Universal Robots PolyScope program: SplitTest.urp

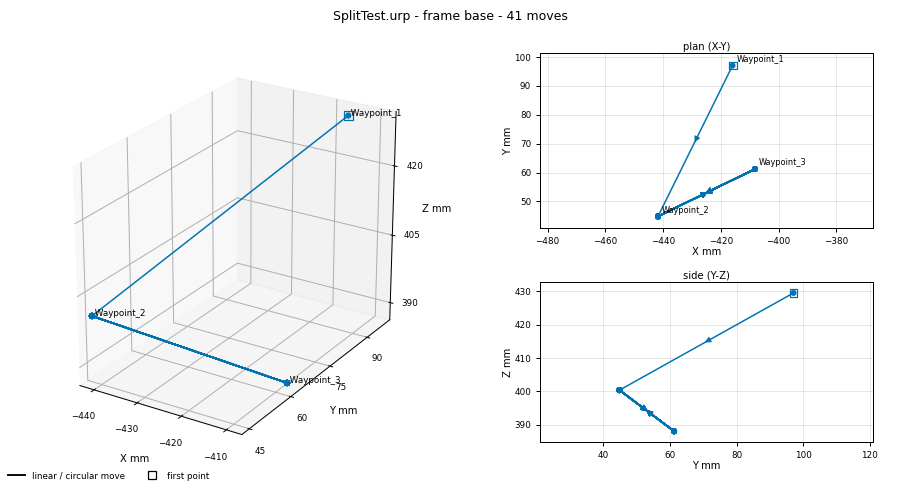
[picture p0: tool path of SplitTest.urp in frame base, 41 of 41 moves have a stored position in this frame; points joined in program order, loops and branches not executed]
Program SplitTest (createdIn=3.0.0 lastSavedIn=3.0.0 directory=/programs installation=default)
Robot Program (runOnlyOnce=true motionType=MoveJ speed=1.047198 acceleration=1.396263 useActiveTCP=false)
  'Program generated by VerticalBot Studio for UR5e on 25/10/2026 12:00:00'
  'Using nominal kinematics.'
  'Using Ref. Frame 2: p[0.100000, -0.050000, 0.020000, 0.000000, 0.000000, 0.523599]'
  'Using TCP Tool 1: p[0.010000, 0.000000, 0.120000, 0.000000, 0.261799, 0.000000]'
  Script: set_tcp(p[0.010000, 0.000000, 0.120000, 0.000000, 0.261799, 0.000000])
  Script: movej([-0.523599, -1.745329, 1.570796, -1.396263, -1.570796, 0.349066],1.20000,0.75000,0,0.0000)
  MoveJ speed 42.97 deg/s, acceleration 68.75 deg/s^2 (useActiveTCP=true)
    Waypoint Waypoint_1: TCP in base x=-415.957 y=97.082 z=429.557 mm, rx=-2.8465 ry=-1.036 rz=-0.3747 rad; joints [-30, -100, 90, -80, -90, 20] deg; flange x=-423.617 y=90.654 z=549.557 mm, rx=2.9521 ry=1.0745 rz=0 rad
  MoveL speed 200 mm/s, acceleration 1200 mm/s^2 (useActiveTCP=true)
    Waypoint Waypoint_2: TCP in base x=-441.769 y=44.852 z=400.392 mm, rx=-2.784 ry=-1.254 rz=-0.442 rad; joints [-22, -96, 90, -80, -90, 20] deg; flange x=-456.215 y=40.554 z=519.861 mm, rx=2.8233 ry=1.257 rz=0.075 rad
    Waypoint Waypoint_3: TCP in base x=-408.198 y=61.237 z=388.074 mm, rx=-2.843 ry=-1.1666 rz=-0.4658 rad; joints [-26, -100, 95, -80, -90, 20] deg; flange x=-424.78 y=58.869 z=507.319 mm, rx=2.8515 ry=1.1521 rz=0.0898 rad
    Waypoint Waypoint_4: TCP in base x=-441.769 y=44.852 z=400.392 mm, rx=-2.784 ry=-1.254 rz=-0.442 rad; joints [-22, -96, 90, -80, -90, 20] deg; flange x=-456.215 y=40.554 z=519.861 mm, rx=2.8233 ry=1.257 rz=0.075 rad
    Waypoint Waypoint_5: TCP in base x=-408.198 y=61.237 z=388.074 mm, rx=-2.843 ry=-1.1666 rz=-0.4658 rad; joints [-26, -100, 95, -80, -90, 20] deg; flange x=-424.78 y=58.869 z=507.319 mm, rx=2.8515 ry=1.1521 rz=0.0898 rad
    Waypoint Waypoint_6: TCP in base x=-441.769 y=44.852 z=400.392 mm, rx=-2.784 ry=-1.254 rz=-0.442 rad; joints [-22, -96, 90, -80, -90, 20] deg; flange x=-456.215 y=40.554 z=519.861 mm, rx=2.8233 ry=1.257 rz=0.075 rad
    Waypoint Waypoint_7: TCP in base x=-408.198 y=61.237 z=388.074 mm, rx=-2.843 ry=-1.1666 rz=-0.4658 rad; joints [-26, -100, 95, -80, -90, 20] deg; flange x=-424.78 y=58.869 z=507.319 mm, rx=2.8515 ry=1.1521 rz=0.0898 rad
    Waypoint Waypoint_8: TCP in base x=-441.769 y=44.852 z=400.392 mm, rx=-2.784 ry=-1.254 rz=-0.442 rad; joints [-22, -96, 90, -80, -90, 20] deg; flange x=-456.215 y=40.554 z=519.861 mm, rx=2.8233 ry=1.257 rz=0.075 rad
    Waypoint Waypoint_9: TCP in base x=-408.198 y=61.237 z=388.074 mm, rx=-2.843 ry=-1.1666 rz=-0.4658 rad; joints [-26, -100, 95, -80, -90, 20] deg; flange x=-424.78 y=58.869 z=507.319 mm, rx=2.8515 ry=1.1521 rz=0.0898 rad
    Waypoint Waypoint_10: TCP in base x=-441.769 y=44.852 z=400.392 mm, rx=-2.784 ry=-1.254 rz=-0.442 rad; joints [-22, -96, 90, -80, -90, 20] deg; flange x=-456.215 y=40.554 z=519.861 mm, rx=2.8233 ry=1.257 rz=0.075 rad
    Waypoint Waypoint_11: TCP in base x=-408.198 y=61.237 z=388.074 mm, rx=-2.843 ry=-1.1666 rz=-0.4658 rad; joints [-26, -100, 95, -80, -90, 20] deg; flange x=-424.78 y=58.869 z=507.319 mm, rx=2.8515 ry=1.1521 rz=0.0898 rad
    Waypoint Waypoint_12: TCP in base x=-441.769 y=44.852 z=400.392 mm, rx=-2.784 ry=-1.254 rz=-0.442 rad; joints [-22, -96, 90, -80, -90, 20] deg; flange x=-456.215 y=40.554 z=519.861 mm, rx=2.8233 ry=1.257 rz=0.075 rad
    Waypoint Waypoint_13: TCP in base x=-408.198 y=61.237 z=388.074 mm, rx=-2.843 ry=-1.1666 rz=-0.4658 rad; joints [-26, -100, 95, -80, -90, 20] deg; flange x=-424.78 y=58.869 z=507.319 mm, rx=2.8515 ry=1.1521 rz=0.0898 rad
    Waypoint Waypoint_14: TCP in base x=-441.769 y=44.852 z=400.392 mm, rx=-2.784 ry=-1.254 rz=-0.442 rad; joints [-22, -96, 90, -80, -90, 20] deg; flange x=-456.215 y=40.554 z=519.861 mm, rx=2.8233 ry=1.257 rz=0.075 rad
    Waypoint Waypoint_15: TCP in base x=-408.198 y=61.237 z=388.074 mm, rx=-2.843 ry=-1.1666 rz=-0.4658 rad; joints [-26, -100, 95, -80, -90, 20] deg; flange x=-424.78 y=58.869 z=507.319 mm, rx=2.8515 ry=1.1521 rz=0.0898 rad
    Waypoint Waypoint_16: TCP in base x=-441.769 y=44.852 z=400.392 mm, rx=-2.784 ry=-1.254 rz=-0.442 rad; joints [-22, -96, 90, -80, -90, 20] deg; flange x=-456.215 y=40.554 z=519.861 mm, rx=2.8233 ry=1.257 rz=0.075 rad
    Waypoint Waypoint_17: TCP in base x=-408.198 y=61.237 z=388.074 mm, rx=-2.843 ry=-1.1666 rz=-0.4658 rad; joints [-26, -100, 95, -80, -90, 20] deg; flange x=-424.78 y=58.869 z=507.319 mm, rx=2.8515 ry=1.1521 rz=0.0898 rad
    Waypoint Waypoint_18: TCP in base x=-441.769 y=44.852 z=400.392 mm, rx=-2.784 ry=-1.254 rz=-0.442 rad; joints [-22, -96, 90, -80, -90, 20] deg; flange x=-456.215 y=40.554 z=519.861 mm, rx=2.8233 ry=1.257 rz=0.075 rad
    Waypoint Waypoint_19: TCP in base x=-408.198 y=61.237 z=388.074 mm, rx=-2.843 ry=-1.1666 rz=-0.4658 rad; joints [-26, -100, 95, -80, -90, 20] deg; flange x=-424.78 y=58.869 z=507.319 mm, rx=2.8515 ry=1.1521 rz=0.0898 rad
    Waypoint Waypoint_20: TCP in base x=-441.769 y=44.852 z=400.392 mm, rx=-2.784 ry=-1.254 rz=-0.442 rad; joints [-22, -96, 90, -80, -90, 20] deg; flange x=-456.215 y=40.554 z=519.861 mm, rx=2.8233 ry=1.257 rz=0.075 rad
    Waypoint Waypoint_21: TCP in base x=-408.198 y=61.237 z=388.074 mm, rx=-2.843 ry=-1.1666 rz=-0.4658 rad; joints [-26, -100, 95, -80, -90, 20] deg; flange x=-424.78 y=58.869 z=507.319 mm, rx=2.8515 ry=1.1521 rz=0.0898 rad
    Waypoint Waypoint_22: TCP in base x=-441.769 y=44.852 z=400.392 mm, rx=-2.784 ry=-1.254 rz=-0.442 rad; joints [-22, -96, 90, -80, -90, 20] deg; flange x=-456.215 y=40.554 z=519.861 mm, rx=2.8233 ry=1.257 rz=0.075 rad
    Waypoint Waypoint_23: TCP in base x=-408.198 y=61.237 z=388.074 mm, rx=-2.843 ry=-1.1666 rz=-0.4658 rad; joints [-26, -100, 95, -80, -90, 20] deg; flange x=-424.78 y=58.869 z=507.319 mm, rx=2.8515 ry=1.1521 rz=0.0898 rad
    Waypoint Waypoint_24: TCP in base x=-441.769 y=44.852 z=400.392 mm, rx=-2.784 ry=-1.254 rz=-0.442 rad; joints [-22, -96, 90, -80, -90, 20] deg; flange x=-456.215 y=40.554 z=519.861 mm, rx=2.8233 ry=1.257 rz=0.075 rad
    Waypoint Waypoint_25: TCP in base x=-408.198 y=61.237 z=388.074 mm, rx=-2.843 ry=-1.1666 rz=-0.4658 rad; joints [-26, -100, 95, -80, -90, 20] deg; flange x=-424.78 y=58.869 z=507.319 mm, rx=2.8515 ry=1.1521 rz=0.0898 rad
    Waypoint Waypoint_26: TCP in base x=-441.769 y=44.852 z=400.392 mm, rx=-2.784 ry=-1.254 rz=-0.442 rad; joints [-22, -96, 90, -80, -90, 20] deg; flange x=-456.215 y=40.554 z=519.861 mm, rx=2.8233 ry=1.257 rz=0.075 rad
    Waypoint Waypoint_27: TCP in base x=-408.198 y=61.237 z=388.074 mm, rx=-2.843 ry=-1.1666 rz=-0.4658 rad; joints [-26, -100, 95, -80, -90, 20] deg; flange x=-424.78 y=58.869 z=507.319 mm, rx=2.8515 ry=1.1521 rz=0.0898 rad
    Waypoint Waypoint_28: TCP in base x=-441.769 y=44.852 z=400.392 mm, rx=-2.784 ry=-1.254 rz=-0.442 rad; joints [-22, -96, 90, -80, -90, 20] deg; flange x=-456.215 y=40.554 z=519.861 mm, rx=2.8233 ry=1.257 rz=0.075 rad
    Waypoint Waypoint_29: TCP in base x=-408.198 y=61.237 z=388.074 mm, rx=-2.843 ry=-1.1666 rz=-0.4658 rad; joints [-26, -100, 95, -80, -90, 20] deg; flange x=-424.78 y=58.869 z=507.319 mm, rx=2.8515 ry=1.1521 rz=0.0898 rad
    Waypoint Waypoint_30: TCP in base x=-441.769 y=44.852 z=400.392 mm, rx=-2.784 ry=-1.254 rz=-0.442 rad; joints [-22, -96, 90, -80, -90, 20] deg; flange x=-456.215 y=40.554 z=519.861 mm, rx=2.8233 ry=1.257 rz=0.075 rad
    Waypoint Waypoint_31: TCP in base x=-408.198 y=61.237 z=388.074 mm, rx=-2.843 ry=-1.1666 rz=-0.4658 rad; joints [-26, -100, 95, -80, -90, 20] deg; flange x=-424.78 y=58.869 z=507.319 mm, rx=2.8515 ry=1.1521 rz=0.0898 rad
    Waypoint Waypoint_32: TCP in base x=-441.769 y=44.852 z=400.392 mm, rx=-2.784 ry=-1.254 rz=-0.442 rad; joints [-22, -96, 90, -80, -90, 20] deg; flange x=-456.215 y=40.554 z=519.861 mm, rx=2.8233 ry=1.257 rz=0.075 rad
    Waypoint Waypoint_33: TCP in base x=-408.198 y=61.237 z=388.074 mm, rx=-2.843 ry=-1.1666 rz=-0.4658 rad; joints [-26, -100, 95, -80, -90, 20] deg; flange x=-424.78 y=58.869 z=507.319 mm, rx=2.8515 ry=1.1521 rz=0.0898 rad
    Waypoint Waypoint_34: TCP in base x=-441.769 y=44.852 z=400.392 mm, rx=-2.784 ry=-1.254 rz=-0.442 rad; joints [-22, -96, 90, -80, -90, 20] deg; flange x=-456.215 y=40.554 z=519.861 mm, rx=2.8233 ry=1.257 rz=0.075 rad
    Waypoint Waypoint_35: TCP in base x=-408.198 y=61.237 z=388.074 mm, rx=-2.843 ry=-1.1666 rz=-0.4658 rad; joints [-26, -100, 95, -80, -90, 20] deg; flange x=-424.78 y=58.869 z=507.319 mm, rx=2.8515 ry=1.1521 rz=0.0898 rad
    Waypoint Waypoint_36: TCP in base x=-441.769 y=44.852 z=400.392 mm, rx=-2.784 ry=-1.254 rz=-0.442 rad; joints [-22, -96, 90, -80, -90, 20] deg; flange x=-456.215 y=40.554 z=519.861 mm, rx=2.8233 ry=1.257 rz=0.075 rad
    Waypoint Waypoint_37: TCP in base x=-408.198 y=61.237 z=388.074 mm, rx=-2.843 ry=-1.1666 rz=-0.4658 rad; joints [-26, -100, 95, -80, -90, 20] deg; flange x=-424.78 y=58.869 z=507.319 mm, rx=2.8515 ry=1.1521 rz=0.0898 rad
    Waypoint Waypoint_38: TCP in base x=-441.769 y=44.852 z=400.392 mm, rx=-2.784 ry=-1.254 rz=-0.442 rad; joints [-22, -96, 90, -80, -90, 20] deg; flange x=-456.215 y=40.554 z=519.861 mm, rx=2.8233 ry=1.257 rz=0.075 rad
    Waypoint Waypoint_39: TCP in base x=-408.198 y=61.237 z=388.074 mm, rx=-2.843 ry=-1.1666 rz=-0.4658 rad; joints [-26, -100, 95, -80, -90, 20] deg; flange x=-424.78 y=58.869 z=507.319 mm, rx=2.8515 ry=1.1521 rz=0.0898 rad
    Waypoint Waypoint_40: TCP in base x=-441.769 y=44.852 z=400.392 mm, rx=-2.784 ry=-1.254 rz=-0.442 rad; joints [-22, -96, 90, -80, -90, 20] deg; flange x=-456.215 y=40.554 z=519.861 mm, rx=2.8233 ry=1.257 rz=0.075 rad
    Waypoint Waypoint_41: TCP in base x=-408.198 y=61.237 z=388.074 mm, rx=-2.843 ry=-1.1666 rz=-0.4658 rad; joints [-26, -100, 95, -80, -90, 20] deg; flange x=-424.78 y=58.869 z=507.319 mm, rx=2.8515 ry=1.1521 rz=0.0898 rad
